// TIA Portal V21 export
// export: Created 2026-08-21T20:18:51.4655298Z, ExportSetting None, DisplayName Totally Integrated Automation Portal, DisplayVersion V21, DisplayName STEP 7 Professional, DisplayVersion V21, DisplayName STEP 7 Safety, DisplayVersion V21, DisplayName Tech WebApplication, DisplayVersion V21, DisplayName WinCC Basic/Comfort/Advanced, DisplayVersion V21, DisplayName WinCC Professional, DisplayVersion V21, DisplayName WinCC Unified, DisplayVersion V21
DATA_BLOCK "Volumeflow_DB"   // DB43
// stored: InstanceOfName Volumeflow, InstanceOfType FB
"Volumeflow"
   // VAR_INPUT
   //    Enable : Bool;
   //    Release_Spd : Int;
   //    T_Release : Real;
   //    Raw_Scale { ExternalAccessible := 'False'; ExternalVisible := 'False'; ExternalWritable := 'False'} : "ScaVal_Raw";
   // END_VAR
   // VAR_OUTPUT
   //    Liter : Real;
   //    Liters_Raw : Int;
   // END_VAR
   // VAR
   //    pi : Real;
   //    r : Real;
   // END_VAR
BEGIN
END_DATA_BLOCK
